Staubli VAL3: simulate.dtx

mdesc mNomSpeed
mdesc mSimulate = {accel=64, vel=80, decel=64, blend=off}
string sMsg
bool bCancel
